(* IEC 61131-3 sources: Lasal-MCP/examples/SampleSource/4_PumpControlSchemeSolution/Stations/MachineControl/MachineControl/Class/VaranManagerPostScan, 1 file *)

(* ---- VaranManagerPostScan.st ---- *)
(*!
<Class
	Name               = "VaranManagerPostScan"
	Revision           = "1.2"
	RealtimeTask       = "false"
	CyclicTask         = "false"
	BackgroundTask     = "false"
	Sigmatek           = "true"
	OSInterface        = "false"
	HighPriority       = "false"
	Automatic          = "false"
	UpdateMode         = "Postscan"
	IconPath           = ".\Class\Tool.ico"
	SharedCommandTable = "true"
	Objectsize         = "(284,120)">
	<Channels>
		<Server Name="Server0" Visualized="true" Initialize="false" WriteProtected="true" Retentive="false"/>
		<Client Name="ManagerConnect" Required="true" Internal="false"/>
	</Channels>
	<RevDoku>
		<Owner Company="Sigmatek"/>
		<Dokumentation Revision="1.2" Date="27.03.2018" Author="EisMic" Company="Sigmatek" Description="Removed CyWork function of class. CyWork of Varanmanager is now called from HwControl."/>
	</RevDoku>
</Class>
*)
VaranManagerPostScan : CLASS
  //Servers:
	Server0 	: SvrChCmd_DINT;
  //Clients:
	ManagerConnect 	: CltChCmd_VaranManager_Base;
  //Variables:
  //Functions:

	FUNCTION VIRTUAL GLOBAL Init;
  //Tables:
	FUNCTION @STD
		VAR_OUTPUT
			ret_code	: CONFSTATES;
		END_VAR;
	FUNCTION GLOBAL TAB @CT_;
END_CLASS;

#pragma usingLtd VaranManager_Base

FUNCTION VIRTUAL GLOBAL VaranManagerPostScan::Init

  IF _FirstScan THEN

#ifdef HWC_LogInit
    HWC_LogInit();
#endif

#ifdef HWC_LogError
    HWC_LogError(this,"@018B (VaranManagerPostScan::Init) Object of VaranManagerPostScan is not used! Cywork of Varanmanager is called by HwControl");
#endif
  END_IF;

END_FUNCTION
